(* IEC 61131-3 sources: RootPLC/conformance/cases/tasks-config, 8 files *)

(* ---- warn_external.st ---- *)
(* spec: [config.external] [scope.vendor-forms]
   expect: warning RP0134
   run: PRG_Main cycles=2
   assert: seen = 4 *)
VAR_GLOBAL
    total : INT;
END_VAR

FUNCTION_BLOCK FB_Add
VAR_EXTERNAL
    total : INT;
END_VAR
total := total + 1;
END_FUNCTION_BLOCK

PROGRAM PRG_Main
VAR
    a, b : FB_Add;
    seen : INT;
END_VAR
a();
b();
seen := total;
END_PROGRAM

(* ---- err_config_unknown_program.st ---- *)
(* spec: [config.program-instance]
   expect: error RP0203 *)
PROGRAM PRG_Main
END_PROGRAM

CONFIGURATION Cfg
    TASK Fast(INTERVAL := T#10ms);
    PROGRAM Main WITH Fast : PRG_Missing;
END_CONFIGURATION

(* ---- err_duplicate_global.st ---- *)
(* spec: [config.global-list]
   expect: error RP0204 *)
CONFIGURATION Cfg
    VAR_GLOBAL
        level : INT;
        level : REAL;
    END_VAR
    RESOURCE Res ON PLC
        TASK Main (INTERVAL := T#10ms, PRIORITY := 1);
        PROGRAM Inst WITH Main : PRG_Main;
    END_RESOURCE
END_CONFIGURATION

PROGRAM PRG_Main
END_PROGRAM

(* ---- ok_configuration.st ---- *)
(* spec: [config.configuration]
   expect: ok
   run: PRG_Main cycles=2
   assert: n = 2 *)
PROGRAM PRG_Main
VAR
    n : INT;
END_VAR
n := n + 1;
END_PROGRAM

CONFIGURATION Cfg
    VAR_GLOBAL
        mode : INT := 1;
    END_VAR
    RESOURCE Res ON PLC
        TASK Fast(INTERVAL := T#10ms, PRIORITY := 1);
        PROGRAM Main WITH Fast : PRG_Main;
    END_RESOURCE
END_CONFIGURATION

(* ---- ok_task.st ---- *)
(* spec: [config.task]
   expect: ok
   run: PRG_Main cycles=1
   assert: n = 1 *)
PROGRAM PRG_Main
VAR
    n : INT;
END_VAR
n := n + 1;
END_PROGRAM

CONFIGURATION Cfg
    RESOURCE Res ON PLC
        TASK Slow(INTERVAL := T#100ms, PRIORITY := 5);
        TASK Fast(INTERVAL := T#1ms);
        PROGRAM Main WITH Fast : PRG_Main;
        PROGRAM Other WITH Slow : PRG_Main;
    END_RESOURCE
END_CONFIGURATION

(* ---- ok_var_config.st ---- *)
(* spec: [config.var-config]
   expect: ok *)
PROGRAM PRG_Main
VAR
    start : BOOL;
END_VAR
END_PROGRAM

CONFIGURATION Cfg
    VAR_CONFIG
        Main.start AT %IX0.0 : BOOL;
    END_VAR
    RESOURCE Res ON PLC
        TASK Fast(INTERVAL := T#10ms);
        PROGRAM Main WITH Fast : PRG_Main;
    END_RESOURCE
END_CONFIGURATION

(* ---- warn_global_list.st ---- *)
(* spec: [config.global-list] [scope.vendor-forms]
   expect: warning RP0134
   run: PRG_Main cycles=3
   assert: c = 13
   assert: last = 13 *)
VAR_GLOBAL CONSTANT
    N_MAX : INT := 3;
    N_LAST : INT := N_MAX + 1;
END_VAR
VAR_GLOBAL
    counter : INT := 10;
    buf : ARRAY[1..N_LAST] OF INT;
END_VAR

PROGRAM PRG_Main
VAR
    last, c : INT;
END_VAR
counter := counter + 1;
buf[N_LAST] := counter;
last := buf[4];
c := counter;
END_PROGRAM

(* ---- warn_globals_per_namespace.st ---- *)
(* spec: [config.global-list] [scope.vendor-forms]
   expect: warning RP0134
   run: PRG_Main cycles=1
   assert: a = 1
   assert: b = 2 *)
NAMESPACE GVL_A
VAR_GLOBAL
    station : INT := 1;
END_VAR
END_NAMESPACE

NAMESPACE GVL_B
VAR_GLOBAL
    station : INT := 2;
END_VAR
END_NAMESPACE

PROGRAM PRG_Main
VAR
    a, b : INT;
END_VAR
a := GVL_A.station;
b := GVL_B.station;
END_PROGRAM
